FUNCTION_BLOCK FB_DomeIdleState EXTENDS  FB_DomeState

VAR
	Stage		: UINT:= 0;
	tonSleep	: TON := (PT:=T#5S);
	tonTimeout	: TON:= (PT:=T#3M); // see Baader Handbook
	tonDelay	: TON:= (PT:=T#20MS);
	
	sSeperator		: STRING := 'd#azi';
	sLeft			: STRING;
	sAzi			: STRING;
	fAzi			: LREAL;
	fAzi_Old		: LREAL;
	// #202: two azimuth readings closer than this (deg) are the same position: the dome reports tenths of a degree
	// and a single step of jitter must not keep the rotation state at slewing (dome_close is refused while slewing)
	fAziTolerance	: LREAL := 0.5;
	bSplitSuccess 	: BOOL;
	
END_VAR


METHOD CloseCommand : BOOL
IF pDome^._DomeRotationState <> E_DomeRotationState.slewing THEN
	Stage:= 0;
	tonSleep(IN:=FALSE);
	tonTimeout(IN:=FALSE);
	tonDelay(IN:=FALSE);
	pDome^.SetState(pDome^.fbDomeCloseingState);
ELSE
	// #202: not silently. The rotation state is slewing as long as two azimuth readings differ.
	LogIgnored(sCommand := 'close (dome rotating)', sLevel := 'WARNING');
END_IF
END_METHOD


METHOD FoundError : BOOL
Stage:= 0;
tonSleep(IN:=FALSE);
tonTimeout(IN:=FALSE);
tonDelay(IN:=FALSE);
pDome^._Error := TRUE;
pDome^.SetState(pDome^.fbDomeErrorState);
END_METHOD

METHOD MoveCommand : BOOL
Stage:= 0;
tonSleep(IN:=FALSE);
tonTimeout(IN:=FALSE);
tonDelay(IN:=FALSE);
pDome^.SetState(pDome^.fbDomeMovingState);
END_METHOD


METHOD OpenCommand : BOOL
Stage:= 0;
tonSleep(IN:=FALSE);
tonTimeout(IN:=FALSE);
tonDelay(IN:=FALSE);
pDome^.SetState(pDome^.fbDomeOpeningState);
END_METHOD


METHOD ParkCommand : BOOL
Stage:= 0;
tonSleep(IN:=FALSE);
tonTimeout(IN:=FALSE);
tonDelay(IN:=FALSE);
pDome^.SetState(pDome^.fbDomeParkingState);
END_METHOD

METHOD RunState : BOOL
VAR_INPUT
END_VAR
// send 'd#getshut' wait for answer
// wait 5 seconds
// send 'd#getazi' wait for answer
CASE Stage OF
	0:
		tonTimeout(IN:=TRUE);
		Stage := 1;
	1:
		pDome^.fbSend(	SendString:= 'd#getshut',
						TXbuffer:= TxBufferDome,
						Busy=>,
						Error=> );
		IF NOT pDome^.fbSend.Busy  THEN
			Stage := 2;
		END_IF
	2: 
		IF pDome^.bStringReceived THEN
			IF pDome^._ReceivedString = 'd#comerro' OR pDome^._ReceivedString = 'd#domerro' THEN
				FoundError();
			ELSIF pDome^._ReceivedString = 'd#shutclo' THEN
				pDome^._DomeShutterState := E_RoofState.closed;
				Stage := 3;
			ELSIF pDome^._ReceivedString = 'd#shutope' THEN
				pDome^._DomeShutterState := E_RoofState.opened;
				Stage := 3;
			ELSIF pDome^._ReceivedString = 'd#shutrun' THEN
				pDome^._DomeShutterState := E_RoofState.unknown;
				Stage := 3;
			END_IF
		ELSIF NOT pDome^.fbReceive.Busy THEN
			tonSleep(IN:=TRUE);
			IF tonSleep.Q THEN
				tonSleep(IN:=FALSE);
				Stage := 1;
			END_IF
		END_IF
		tonTimeout(IN:=TRUE);
		IF tonTimeout.Q THEN
			tonTimeout(IN:=FALSE);
			FoundError();
		END_IF
	3:
		tonTimeout(IN:=FALSE);
		tonSleep(IN:=TRUE);
		IF tonSleep.Q THEN
			tonSleep(IN:=FALSE);
			Stage := 4;
			tonTimeout(IN:=TRUE);
		END_IF
	4:
		pDome^.fbSend(	SendString:= 'd#getazim',
						TXbuffer:= TxBufferDome,
						Busy=>,
						Error=> );
		IF NOT pDome^.fbSend.Busy  THEN
			Stage := 5;
		END_IF
	5: 
		IF pDome^._HasReceivedString THEN
			IF pDome^._ReceivedString = 'd#comerro' OR pDome^._ReceivedString = 'd#domerro' THEN
				FoundError();
			ELSE
				bSplitSuccess := FindAndSplit(
									pSeparator := ADR(sSeperator),
									pSrcString := ADR(pDome^.sReceivedString),
									pLeftString:= ADR(sLeft),
									nLeftSize	:= 1,
									pRightString := ADR(sAzi),
									nRightSize := 5,
									bSearchFromRight:= FALSE);
									
				IF bSplitSuccess AND ( STRING_TO_LREAL(sAzi) <> 0 OR sAzi = '0000') THEN
					// (STRING_TO_LREAL(sAzi) <> 0 OR sAzi := '0000') -> either sAzi actual 0 OR STRING_TO_LREAL error
					fAzi := STRING_TO_LREAL(sAzi)/10.0;
					//Baader measures azimuth as West of South, so we need to convert it. This works both ways.
					IF fAzi  >= 180.0 THEN
						pDome^._Position := fAzi - 180.0;
					ELSE
						pDome^._Position := fAzi + 180.0;
					END_IF
					IF ABS(fAzi - fAzi_Old) < fAziTolerance THEN
						IF ABS(pDome^.Position - 180.0) < 5.0 THEN
							pDome^._DomeRotationState := E_DomeRotationState.parked;
						ELSE
							pDome^._DomeRotationState := E_DomeRotationState.idle;
						END_IF
					ELSE
						pDome^._DomeRotationState := E_DomeRotationState.slewing;
					END_IF
					fAzi_Old := fAzi;
					Stage := 6;
				END_IF
			END_IF
		ELSIF NOT pDome^.fbReceive.Busy THEN
			tonSleep(IN:=TRUE);
			IF tonSleep.Q THEN
				tonSleep(IN:=FALSE);
				Stage := 4;
			END_IF
		END_IF
		tonTimeout(IN:=TRUE);
		IF tonTimeout.Q THEN
			tonTimeout(IN:=FALSE);
			FoundError();
		END_IF
	6:
		tonTimeout(IN:=FALSE);
		IF ABS( pDome^.Position - pDome^._Position) > 10.0 AND pDome^._Track THEN
			MoveCommand();
		ELSE
			Stage:= 7;
		END_IF
	7:
		tonSleep(IN:=TRUE);
		IF tonSleep.Q THEN
			tonSleep(IN:=FALSE);
			Stage := 0;
		END_IF		
END_CASE
END_METHOD


METHOD StopCommand : BOOL
Stage:= 0;
tonSleep(IN:=FALSE);
tonTimeout(IN:=FALSE);
tonDelay(IN:=FALSE);
pDome^.SetState(pDome^.fbDomeStoppingState);
END_METHOD


PROPERTY StateID : STRING
GET
StateID := 'Idle State';
END_GET
END_PROPERTY

END_FUNCTION_BLOCK

(* stored: Version 1.1.0.1, ProductVersion 3.1.4024.15
   POU FB_DomeIdleState: Id {18941870-4fd2-48dc-9e55-0c95299f7dd7}, SpecialFunc None
   Method CloseCommand: Id {672045a5-18c7-44e8-b963-3dfd226f80ee}
   Method FoundError: Id {b1011a7e-754f-4d17-83aa-eb0986f7d112}
   Method MoveCommand: Id {f3c4f054-a43b-464f-8284-7288eb1f1cb3}
   Method OpenCommand: Id {336403ce-c239-42a6-9c74-883457eb74c5}
   Method ParkCommand: Id {87d7fae6-5a44-4333-ac1f-722c8d011ed6}
   Method RunState: Id {cb13016a-e3a1-402f-bad4-fdf6a2718530}
   Method StopCommand: Id {7acaa647-1f4d-457c-aae9-b2517072faf9}
   Property StateID: Id {25716fec-f7ae-4751-8f4c-4e9b44cfd178}
   Get Get: Id {51112923-8420-482a-8c35-1fc4b0cd957c} *)
